(*
SPDX-FileCopyrightText: © 2026 Oleksandr Tiutyk <trofimich@gmail.com>
SPDX-License-Identifier: MIT
License: https://opensource.org/license/mit
*)

(*!
<summary>Orders DATE_AND_TIME values described by generic descriptors.</summary>
<description>
Non-null addresses must reference live DATE_AND_TIME storage. TypeClass and Size are not validated and no
numeric conversion is performed. Two null addresses compare equal; one null address sorts before a non-null
address. Descriptors are passed by value; payload remains borrowed and is not modified, cloned, released or
retained. IsMemoryOwner does not affect comparison.
</description>
*)

FUNCTION_BLOCK DateAndTimeComparer EXTENDS TOF_Core.Object IMPLEMENTS TOF_Core.IComparer
VAR_STAT
	//! <summary>Class name shared by all instances of this function block.</summary>
	{attribute 'hide'} 
	_ClassName : STRING := __POUNAME();
END_VAR

{attribute 'monitoring' := 'call'}
PROPERTY ClassName : REFERENCE TO STRING
GET
ClassName REF= _ClassName;
END_GET
END_PROPERTY

(*!
<summary>Compares the first operand with the second using this ordering strategy.</summary>
<description>
Non-null addresses must reference live DATE_AND_TIME storage. TypeClass and Size are not validated and no
numeric conversion is performed. Two null addresses compare equal; one null address sorts before a non-null
address. Descriptors are passed by value; payload remains borrowed and is not modified, cloned, released or
retained. IsMemoryOwner does not affect comparison. Descendants cannot replace this standard ordering;
implement IComparer separately for a different ordering strategy.
</description>
*)
//!<param name="first">First descriptor; referenced storage is borrowed for the call.</param>
//!<param name="second">Second descriptor; referenced storage is borrowed for the call.</param>
{attribute "object_name" := "Compare"}
METHOD FINAL Compare : TOF_Core.COMPARISON_RESULT
VAR_INPUT
	first : TOF_Core.GENERIC_VALUE;
	second : TOF_Core.GENERIC_VALUE;
END_VAR
VAR
	leftPointer : POINTER TO DATE_AND_TIME; 
	rightPointer : POINTER TO DATE_AND_TIME; 
END_VAR
IF first.Address = 0 AND_THEN second.Address = 0 THEN
	Compare := TOF_Core.COMPARISON_RESULT.FIRST_EQUAL_TO_SECOND;
	RETURN;
END_IF

IF first.Address = 0 THEN
	Compare := TOF_Core.COMPARISON_RESULT.FIRST_LESS_THAN_SECOND;
	RETURN;	
END_IF

IF second.Address = 0 THEN
	Compare := TOF_Core.COMPARISON_RESULT.FIRST_GREATER_THAN_SECOND;
	RETURN;	
END_IF

leftPointer := first.Address;
rightPointer := second.Address;

IF leftPointer^ < rightPointer^ THEN
	Compare := TOF_Core.COMPARISON_RESULT.FIRST_LESS_THAN_SECOND;
ELSIF leftPointer^ > rightPointer^ THEN
	Compare := TOF_Core.COMPARISON_RESULT.FIRST_GREATER_THAN_SECOND;
ELSE
	Compare := TOF_Core.COMPARISON_RESULT.FIRST_EQUAL_TO_SECOND;	
END_IF
END_METHOD

{attribute 'monitoring' := 'call'}
PROPERTY NamespaceName : REFERENCE TO STRING
GET
NamespaceName REF= CurrentNamespace.Name;
END_GET
END_PROPERTY

{attribute 'monitoring' := 'call'}
PROPERTY SelfSize : ULINT
GET
SelfSize := XSIZEOF(THIS^);
END_GET
END_PROPERTY

END_FUNCTION_BLOCK

(* stored: Version 1.1.0.1
   POU DateAndTimeComparer: Id {c7624954-7866-4335-b6ea-542bbc0f5ff3}, SpecialFunc None
   Property ClassName: Id {c7158c9a-41c2-4bf7-b154-cda0e5f6fe61}
   Get Get: Id {3cf85dee-d11d-4346-a9bd-dcb2db67323b}
   Method Compare: Id {5fa917ff-f4ed-433b-afa5-de1963f626e1}
   Property NamespaceName: Id {1ec9f00a-cc70-4a3c-8c23-ca9da2e44002}
   Get Get: Id {8e3bb480-4398-4f13-9eba-3ac20a70921a}
   Property SelfSize: Id {b6e75391-1b1f-46f9-9a33-6f5c36086d2b}
   Get Get: Id {ca34781c-13ed-4e6c-a3d9-106c7d41417a} *)
